(*
SPDX-FileCopyrightText: c 2026 Oleksandr Tiutyk <trofimich@gmail.com>
SPDX-License-Identifier: MIT
License: https://opensource.org/license/mit
*)

(*!
<summary>Checks fitted concatenation, including the 255-character boundary.</summary>
<description>
Uses one task and stays at a stable address while assertions are bound to this instance.
</description>
*)

{attribute 'no_assign'}
{attribute 'no_explicit_call' := 'do not call this function block directly'}
FUNCTION_BLOCK StringConcatFitTest EXTENDS TOF_Testing.SingleCycleTest
VAR_STAT
	{attribute 'hide'}
	_ClassName : STRING := __POUNAME();
END_VAR

(*!
<summary>Checks fitted concatenation, including the 255-character boundary.</summary>
<description>
Distinct ASCII fragments reveal the first discarded byte and any changes in fragment order. Compares all
255 bytes against a separately assembled expected result.
</description>
*)
METHOD PROTECTED ExecuteTest
VAR
	text : STRING(255);
	first : STRING(100) := 'aaaaaaaaaaaaaaaaaaaaaaaaaaaaaaaaaaaaaaaaaaaaaaaaaaaaaaaaaaaaaaaaaaaaaaaaaaaaaaaaaaaaaaaaaaaaaaaaaaaa';
	second : STRING(100) := 'bbbbbbbbbbbbbbbbbbbbbbbbbbbbbbbbbbbbbbbbbbbbbbbbbbbbbbbbbbbbbbbbbbbbbbbbbbbbbbbbbbbbbbbbbbbbbbbbbbbb';
	third : STRING(100) := 'cccccccccccccccccccccccccccccccccccccccccccccccccccccccccccccccccccccccccccccccccccccccccccccccccccc';
	expectedText : STRING(255);
END_VAR
text := TOF_Core.Strings.ConcatFit255('Hello, ', 'World!');
Assert.ThatBool(
	actual := text = 'Hello, World!',
	message := "ConcatFit255 must preserve an ordinary fit"
).IsTrue();

text := TOF_Core.Strings.ConcatFit255('Part1', '', 'Part2', '', 'Part3');
Assert.ThatBool(
	actual := text = 'Part1Part2Part3',
	message := "ConcatFit255 must skip empty fragments without stopping"
).IsTrue();

text := TOF_Core.Strings.ConcatFit255(first, second, third);
Assert.ThatInt(
	actual := Tc2_Standard.LEN(STR := text),
	message := "ConcatFit255 must fill the 255-character result"
).ToBe(expected := 255);

// The first two 100-byte fragments leave room for 52 bytes from the third and the three-dot suffix.
expectedText := Tc2_Standard.CONCAT(STR1 := first, STR2 := second);
expectedText := Tc2_Standard.CONCAT(
	STR1 := expectedText,
	STR2 := 'cccccccccccccccccccccccccccccccccccccccccccccccccccc...'
);
Assert.ThatBool(
	actual := text = expectedText,
	message := "Truncation must preserve the 252-byte prefix and end in three dots"
).IsTrue();
END_METHOD

//! <summary>Borrows the concrete class name. Callers must not modify it.</summary>
{attribute 'monitoring' := 'call'}
PROPERTY ClassName : REFERENCE TO STRING
GET
ClassName REF= _ClassName;
END_GET
END_PROPERTY

//! <summary>Borrows the compiler-initialized namespace name. Callers must not modify it.</summary>
{attribute 'monitoring' := 'call'}
PROPERTY NamespaceName : REFERENCE TO STRING
GET
NamespaceName REF= CurrentNamespace.Name;
END_GET
END_PROPERTY

//! <summary>Reports the concrete instance size in bytes.</summary>
{attribute 'monitoring' := 'call'}
PROPERTY SelfSize : ULINT
GET
SelfSize := XSIZEOF(THIS^);
END_GET
END_PROPERTY

END_FUNCTION_BLOCK

(* stored: Version 1.1.0.1
   POU StringConcatFitTest: Id {18ffe0bc-42d6-476f-831c-25bf10f6dbc3}, SpecialFunc None
   Method ExecuteTest: Id {c67d781f-01d2-4798-8934-37193315e412}
   Property ClassName: Id {97d366a8-bc7f-43ff-a96e-f3fb4fa9e35d}
   Get Get: Id {01bbef21-c9a3-474e-8099-243de193d9c8}
   Property NamespaceName: Id {6331f5e3-bc02-482c-bc47-e500610d0b2f}
   Get Get: Id {25a18d73-7905-44d6-b074-2d1b280b915e}
   Property SelfSize: Id {b2fa4aee-a63a-4add-bdbd-b625bd94db55}
   Get Get: Id {7cf46a53-4cb4-44e8-a353-1a4e6347b8ba} *)
